(*
SPDX-FileCopyrightText: © 2026 Oleksandr Tiutyk <trofimich@gmail.com>
SPDX-License-Identifier: MIT
License: https://opensource.org/license/mit
*)

(*!
<summary>Reports an argument whose TwinCAT type class is not supported by the operation.</summary>
<description>
The caller detects the invalid argument. Throw records a diagnostic message and source metadata; it does not
inspect the actual argument or decide which types are supported. Dynamic instances belong to the current task
memory manager until cleanup. Dynamic copies are explicitly registered by Clone after construction; plain
__NEW does not transfer ownership to the task manager.
Runtime type diagnostics use TYPE_ names for known classes and decimal codes for unknown values.
</description>
*)

{attribute 'enable_dynamic_creation'}
{attribute 'no_explicit_call' := 'do not call this function block directly'}
FUNCTION_BLOCK ArgumentTypeClassNotSupportedException EXTENDS GeneralException IMPLEMENTS IArgumentTypeClassNotSupportedException
VAR_STAT
	//! <summary>Class name shared by all instances of this function block.</summary>
	{attribute 'hide'} 
	_ClassName : STRING := __POUNAME();
END_VAR

{attribute 'monitoring' := 'call'}
PROPERTY ClassName : REFERENCE TO STRING
GET
ClassName REF= _ClassName;
END_GET
END_PROPERTY

(*!
<summary>Creates a distinct auto-disposed copy of this concrete exception type.</summary>
<description>
Copies message, code, source and timestamps through CopyGeneralFields; any prepared inner cause remains
borrowed. The current task memory manager owns the clone until cleanup. Allocation failure is terminal.
Descendants with additional payload must override Clone to preserve their type and fields. Registers the newly
constructed instance before copying payload, outside FB_init. Registration failure releases the unregistered
instance and raises a terminal error; copy failure leaves the registered instance owned by the task manager
for cleanup. Custom overrides must follow the same ownership sequence.
</description>
*)
METHOD Clone : IObject
VAR
	exceptionClone : POINTER TO ArgumentTypeClassNotSupportedException;
END_VAR
exceptionClone := __NEW(ArgumentTypeClassNotSupportedException);

IF exceptionClone = 0 THEN
	DynamicMemoryManager.RaiseAllocationFailure();
END_IF

DynamicMemoryManager.RegisterAutoDisposedObject(autoDisposedObject := exceptionClone^);

exceptionClone^.CopyGeneralFields(sourceException := THIS^);

Clone := exceptionClone^;
END_METHOD

(*!
<summary>Provides the library namespace used in diagnostics.</summary>
<description>
Borrowed read-only reference to the compiler-initialized library namespace; no ownership transfer.
</description>
*)
{attribute 'monitoring' := 'call'}
PROPERTY NamespaceName : REFERENCE TO STRING
GET
NamespaceName REF= CurrentNamespace.Name;
END_GET
END_PROPERTY

(*!
<summary>Reports the byte size of this concrete instance.</summary>
<description>
Uses XSIZEOF on the instance. Does not include separately allocated payloads or prove that an arbitrary
address is valid.
</description>
*)
{attribute 'monitoring' := 'call'}
PROPERTY SelfSize : ULINT
GET
SelfSize := XSIZEOF(THIS^);
END_GET
END_PROPERTY

(*!
<summary>Builds the argument diagnostic and propagates this exception.</summary>
<description>
Call in the owning cyclic task, not during FB_init. Captures message, source and timestamps with zero error
code and no inner cause. Supplied names are copied into a local buffer without heap allocation; no caller
storage is retained. Exception clone allocation failure follows the shared terminal memory mechanism.
Known runtime type classes appear by their TYPE_ names; unknown values retain their decimal codes.
</description>
<param name="argumentName">Name of the argument rejected by the caller.</param>
*)
METHOD Throw
VAR_INPUT
	sourceNamespaceName : STRING;
	sourceClassName : STRING;
	sourcePOUName : STRING;
	sourcePosition : STRING;
	argumentName : STRING;
	argumentType : __SYSTEM.TYPE_CLASS;
END_VAR
VAR
	message : ERROR_MESSAGE;
END_VAR
WideStrings.Append255(
	message,
	"Argument '",
	TO_WSTRING(argumentName),
	"' has not supported type class '",
	SystemTypeClassConvertor.ToWideString(typeClass := argumentType),
	"' in '",
	TO_WSTRING(GetFullPOUName(
		sourceNamespaceName := sourceNamespaceName,
		sourceClassName := sourceClassName,
		sourcePOUName := sourcePOUName
	)),
	"'");

InternalThrow(
	sourceNamespaceName := sourceNamespaceName,
	sourceClassName := sourceClassName,
	sourcePOUName := sourcePOUName,
	sourcePosition := sourcePosition,
	message := message,
	errorCode := 0,
	innerException := 0
);
END_METHOD

END_FUNCTION_BLOCK

(* stored: Version 1.1.0.1
   POU ArgumentTypeClassNotSupportedException: Id {70be0cc3-2d2a-41e4-a517-12fc32079b0e}, SpecialFunc None
   Property ClassName: Id {b324b57f-066f-4cb6-b0ac-ec9d24afe8c8}
   Get Get: Id {61c7bed7-5023-47b9-86ea-5957a1e30b10}
   Method Clone: Id {46c54889-37ea-46c8-9aa0-acf43a681cd3}
   Property NamespaceName: Id {1f6edfcd-d71b-4a39-907c-8c955c3ee813}
   Get Get: Id {bef4fbcc-f50d-4117-9a43-eccb05a690ef}
   Property SelfSize: Id {e6a7413c-f3e8-4086-8370-46248199af7e}
   Get Get: Id {61d6a2ea-1d21-4076-8c14-7090dd60a922}
   Method Throw: Id {82d8fa01-6199-47ad-8e53-39c23c88c3d9} *)
